Fanuc KAREL source: KT00759.KL

PROGRAM KT00759
%NOLOCKGROUP
VAR
  S1: STRING[80]
  S2: STRING[80]
  OUT: REAL
BEGIN
  S1 = 'A'
  S2 = 'B'
  S1 = 'A'
  S2 = 'B'
  OUT = ABS(S1)
END KT00759
